FUNCTION_BLOCK ARM_IMC (* Extracted Composite Function Block Type *)
  (* Standard: 61499-2 *)
  (* Version 10/27/2026, lizar *)
  PACKAGE Main;
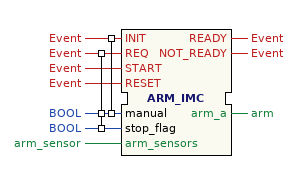
  EVENT_INPUT
    INIT WITH manual; (* Initialization Request *)
    REQ WITH manual, stop_flag; (* Normal Execution Request *)
    START;
    RESET;
  END_EVENT
  EVENT_OUTPUT
    READY;
    NOT_READY;
  END_EVENT
  VAR_INPUT
    manual : BOOL;
    stop_flag : BOOL;
  END_VAR
  SOCKETS
    arm_sensors : arm_sensor;
  END_SOCKETS
  PLUGS
    arm_a : arm;
  END_PLUGS
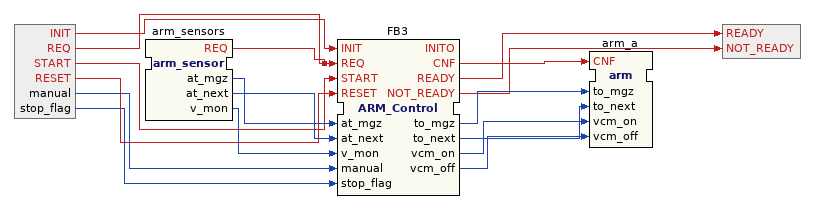
  FBS
    FB3 : ARM_Control;
  END_FBS
  EVENT_CONNECTIONS
    INIT TO FB3.INIT;
    REQ TO FB3.REQ;
    START TO FB3.START;
    RESET TO FB3.RESET;
    FB3.READY TO READY;
    FB3.NOT_READY TO NOT_READY;
    FB3.CNF TO arm_a.CNF;
    arm_sensors.REQ TO FB3.REQ;
  END_CONNECTIONS
  DATA_CONNECTIONS
    manual TO FB3.manual;
    stop_flag TO FB3.stop_flag;
    FB3.to_mgz TO arm_a.to_mgz;
    FB3.to_next TO arm_a.to_next;
    FB3.vcm_on TO arm_a.vcm_on;
    FB3.vcm_off TO arm_a.vcm_off;
    arm_sensors.at_mgz TO FB3.at_mgz;
    arm_sensors.at_next TO FB3.at_next;
    arm_sensors.v_mon TO FB3.v_mon;
  END_CONNECTIONS
END_FUNCTION_BLOCK
